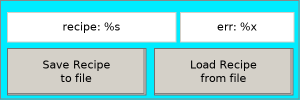
VISUALIZATION vis_RecipeControl_v01  // 300x100
VAR_INPUT
	Definition: STRING;
END_VAR
VAR
	RecipeName: STRING:='name';
END_VAR
    Button (7,48 139x47), "Save Recipe to file"
        OnMouseClick: ExecuteCommand ExecuteCommand=ExecuteCommand=[Command=CreateRecipe, Value=Definition, Value2=RecipeName, Command=SaveRecipeAs, Value=Definition, Value2=RecipeName]
    Button (154,48 139x47), "Load Recipe from file"
        OnMouseClick: ExecuteCommand ExecuteCommand=ExecuteCommand=[Command=LoadRecipeFrom, Value=Definition, Value2=RecipeName]
    Textfield (7,12 169x30), "recipe: %s", text variable: Definition
    Textfield (180,12 114x30), "err: %x", text variable: prg_RecipeManager.LastError, colour toggle: prg_RecipeManager.LastError<>0
        toggle prg_RecipeManager.bResetError
END_VISUALIZATION

(* stored: Version 1.1.0.1, ProductVersion 3.1.4024.12
   Visu vis_RecipeControl_v01: Id {2625c674-a409-41c7-a51b-d401c34acdcc} *)
